Fanuc KAREL source: kb00002.KL

-- PROVISIONAL review KL for V770-1; original PC SHA256 35a25fc0e524ba14f2dbf7950372437b694950c687b8337f64c73d5d55f8e5f6
-- Incomplete behavior may be omitted. Consult companion uncertainty JSON. Do not deploy.
PROGRAM KB00002
%NOLOCKGROUP
VAR
  P1 : INTEGER
  RESULT : INTEGER
BEGIN
  -- UNRESOLVED_PC offsets 5-12; opcodes 9D,23
  -- UNRESOLVED_PC offsets 17-30; opcodes 21,50,23
  -- UNRESOLVED_PC offsets 35-39; opcodes 7F
END KB00002
